Fanuc KAREL source: KT00594.KL

PROGRAM KT00594
%NOLOCKGROUP
VAR
  I1: INTEGER
  R2: REAL
  OUT: STRING[80]
BEGIN
  I1 = 2
    R2 = 3.0
  OUT = I1 + R2
END KT00594
